TYPE ST_VisuXtsGantry :
STRUCT
	(* One visualised XTS gantry (e.g. IDH). Register the instance's symbol path in the manifest with
	   eType := E_VisuComponentType.XTS_GANTRY. *)
	stConfig : ST_VisuXtsGantryConfig; // read at discovery and after nConfigVersion changes
	stState : ST_VisuXtsGantryState; // read every gateway cycle
END_STRUCT
END_TYPE

(* stored: Version 1.1.0.1, ProductVersion 3.1.4026.18
   DUT ST_VisuXtsGantry: Id {4b6fcae5-7e81-4610-9da1-6ce7c703ab41} *)
